// =============================================================================
// s7-to-codesys — корпус SCL. Написан с нуля, объект вымышленный (ВОС «Северная»).
//
// Файл:   FB_Valve.scl
// Блок:   FUNCTION_BLOCK "FB_Valve"
// -----------------------------------------------------------------------------
// Назначение
//   Задвижка с электроприводом (открыть/закрыть, два концевика) с контролем
//   времени хода. Для пилотного бистабильного распределителя дополнительно
//   формируются импульсы pulseOpen/pulseClose. Экземпляр DB_XV201 (подача
//   исходной воды на фильтр).
//
// Логика (нормативное описание)
//   Состояния state: 0 — неизвестно, 1 — закрыта, 2 — открывается, 3 — открыта,
//   4 — закрывается, 9 — авария. Коды faultCode: 1 — не дошла за travelTime,
//   2 — оба концевика одновременно, 3 — самопроизвольный уход с концевика.
//   1. Концевики проходят через мультиэкземпляры "FB_Debounce" (задержки по
//      умолчанию): isOpen, isClosed.
//   2. По фронту reset (R_TRIG), если не оба концевика: state := 0, faultCode := 0.
//   3. Оба концевика (isOpen AND isClosed): state := 9, faultCode := 2 (сразу).
//   4. Таймеры хода: TON_TIME(IN := state = 2, PT := travelTime) и
//      TON_TIME(IN := state = 4, PT := travelTime) — вызываются до переходов.
//      Уход с концевика — спад isOpen / isClosed (F_TRIG).
//   5. Переходы (CASE state, один за вызов):
//        0: cmdClose -> 4; иначе cmdOpen -> 2; иначе isClosed -> 1; иначе isOpen -> 3;
//        1: cmdOpen AND NOT cmdClose -> 2; спад isClosed -> 9 (код 3);
//        2: cmdClose -> 4; isOpen -> 3; таймер открытия -> 9 (код 1);
//        3: cmdClose -> 4; спад isOpen -> 9 (код 3);
//        4: isClosed -> 1; cmdOpen AND NOT cmdClose -> 2; таймер закрытия -> 9 (код 1);
//        9: ожидание сброса; другое значение -> 0.
//   6. coilOpen := state = 2; coilClose := state = 4 (реверсивный пускатель);
//      pulseOpen / pulseClose — TP_TIME длиной pulseTime по входу в состояние 2 / 4.
// Что проверяет при конвертации
//   мультиэкземпляр пользовательского ФБ с типом в кавычках, обращение к его
//   выходу (#debOpen.debounced), TP_TIME, F_TRIG, CASE с несколькими операторами
//   в ветке, метки-литералы.
// =============================================================================
FUNCTION_BLOCK "FB_Valve"
TITLE = Motorized valve with travel monitoring
{ S7_Optimized_Access := 'TRUE' }
AUTHOR : WTP2
FAMILY : Valves
VERSION : 1.2
//Задвижка: команды, концевики, контроль хода
   VAR_INPUT
      cmdOpen : Bool;   // Команда «открыть» (уровень)
      cmdClose : Bool;   // Команда «закрыть» (уровень), приоритет над «открыть»
      limitOpen : Bool;   // Концевик «открыто»
      limitClosed : Bool;   // Концевик «закрыто»
      reset : Bool;   // Сброс аварии (по фронту)
      travelTime : Time := T#30S;   // Предельное время хода
      pulseTime : Time := T#1S;   // Длительность импульса на пилот
   END_VAR

   VAR_OUTPUT
      coilOpen : Bool;   // Пускатель «открыть»
      coilClose : Bool;   // Пускатель «закрыть»
      pulseOpen : Bool;   // Импульс «открыть» на пилот
      pulseClose : Bool;   // Импульс «закрыть» на пилот
      isOpen : Bool;   // Открыта (после фильтра)
      isClosed : Bool;   // Закрыта (после фильтра)
      state : Int;   // Состояние
      faultCode : Int;   // Код аварии
   END_VAR

   VAR
      debOpen : "FB_Debounce";   // Фильтр концевика «открыто»
      debClosed : "FB_Debounce";   // Фильтр концевика «закрыто»
      tonOpening {InstructionName := 'TON_TIME'; LibVersion := '1.0'} : TON_TIME;
      tonClosing {InstructionName := 'TON_TIME'; LibVersion := '1.0'} : TON_TIME;
      tpOpen {InstructionName := 'TP_TIME'; LibVersion := '1.0'} : TP_TIME;
      tpClose {InstructionName := 'TP_TIME'; LibVersion := '1.0'} : TP_TIME;
      edgeReset {InstructionName := 'R_TRIG'; LibVersion := '1.0'} : R_TRIG;
      lostOpen {InstructionName := 'F_TRIG'; LibVersion := '1.0'} : F_TRIG;
      lostClosed {InstructionName := 'F_TRIG'; LibVersion := '1.0'} : F_TRIG;
   END_VAR


BEGIN
    REGION Limit switches
        #debOpen(raw := #limitOpen);
        #debClosed(raw := #limitClosed);
        #isOpen := #debOpen.debounced;
        #isClosed := #debClosed.debounced;
    END_REGION

    REGION Reset and discrepancy
        #edgeReset(CLK := #reset);
        IF #edgeReset.Q AND NOT (#isOpen AND #isClosed) THEN
            #state := 0;
            #faultCode := 0;
        END_IF;
        IF #isOpen AND #isClosed THEN
            #state := 9;
            #faultCode := 2;
        END_IF;
    END_REGION

    REGION State machine
        #tonOpening(IN := #state = 2, PT := #travelTime);
        #tonClosing(IN := #state = 4, PT := #travelTime);
        #lostOpen(CLK := #isOpen);
        #lostClosed(CLK := #isClosed);

        CASE #state OF
            0:
                IF #cmdClose THEN
                    #state := 4;
                ELSIF #cmdOpen THEN
                    #state := 2;
                ELSIF #isClosed THEN
                    #state := 1;
                ELSIF #isOpen THEN
                    #state := 3;
                END_IF;
            1:
                IF #cmdOpen AND NOT #cmdClose THEN
                    #state := 2;
                ELSIF #lostClosed.Q THEN
                    #state := 9;
                    #faultCode := 3;
                END_IF;
            2:
                IF #cmdClose THEN
                    #state := 4;
                ELSIF #isOpen THEN
                    #state := 3;
                ELSIF #tonOpening.Q THEN
                    #state := 9;
                    #faultCode := 1;
                END_IF;
            3:
                IF #cmdClose THEN
                    #state := 4;
                ELSIF #lostOpen.Q THEN
                    #state := 9;
                    #faultCode := 3;
                END_IF;
            4:
                IF #isClosed THEN
                    #state := 1;
                ELSIF #cmdOpen AND NOT #cmdClose THEN
                    #state := 2;
                ELSIF #tonClosing.Q THEN
                    #state := 9;
                    #faultCode := 1;
                END_IF;
            9:
                ;   // ожидание сброса
            ELSE
                #state := 0;
        END_CASE;
    END_REGION

    REGION Outputs
        #coilOpen := #state = 2;
        #coilClose := #state = 4;
        #tpOpen(IN := #state = 2, PT := #pulseTime);
        #tpClose(IN := #state = 4, PT := #pulseTime);
        #pulseOpen := #tpOpen.Q;
        #pulseClose := #tpClose.Q;
    END_REGION

END_FUNCTION_BLOCK

